FUNCTION UINT_TO_E_TablePosition : E_TablePosition
VAR_INPUT
    uiPosition : UINT;
END_VAR

CASE uiPosition OF
    1:
        UINT_TO_E_TablePosition := E_TablePosition.Position1;

    2:
        UINT_TO_E_TablePosition := E_TablePosition.Position2;

    3:
        UINT_TO_E_TablePosition := E_TablePosition.Position3;

    4:
        UINT_TO_E_TablePosition := E_TablePosition.Position4;

ELSE
    UINT_TO_E_TablePosition := E_TablePosition.Unknown;
END_CASE

END_FUNCTION

(* stored: Version 1.1.0.1, ProductVersion 3.1.4026.18
   POU UINT_TO_E_TablePosition: Id {74f1f88a-2b96-4cb9-99c4-c5b6acc10bf1}, SpecialFunc None *)
